(* IEC 61131-3 sources: s7-to-codesys/src/POUs/Lang/Converted/FB_BackwashGraph, 2 files *)

(* ---- FB_BackwashGraph.decl.st ---- *)
// Назначение: Промывка фильтра (GRAPH)
//             Промывка скорого фильтра (GRAPH S7-1500), шаги S1–S6. S1 Idle (начальный): N xReady.
//             T1 Start: xStart. S2 Drain: N xDrainValve, S xWashActive, событие S1 — iWashCount + 1;
//             контроль xValveFault держит шаг до квитирования ACK_EF (ERR_FLT = 1). После S2 альтернатива:
//             T2 LongWash (xLevelLow AND NOT xShortWash) — параллельно S3 Air (N xBlower, D xAirValve 2 с)
//             и S4 Rinse (NC xWashPump, блокировка xPumpOk), синхронизация T4 AirDone: Air.T >= 10 с;
//             T3 ShortWash (xLevelLow AND xShortWash) — S5 QuickRinse (N xWashPump), T5 QuickDone: xLevelHigh.
//             S6 Refill: N xInletValve, R xWashActive; T6 Full: xLevelHigh — прыжок к S1. Постоперация:
//             xValvesBusy := xDrainValve OR xInletValve. INIT_SQ — начальное состояние, OFF_SQ — шаги выключены.
// Автор:      WTP2 (исходный блок S7); перевод в ST — s7conv 0.1.0
// Версия:     0.1 (исходный блок S7)
// Документ:   docs/CONVERSION_REPORT.md, docs/MAPPING.md
// Источник:   samples/lang/FB_BackwashGraph.xml, GRAPH, SW.Blocks.FB "FB_BackwashGraph", пространство имён
//             Interface/v5, FAMILY Filters
// Сгенерировано s7conv: пометки MIGRATION-CHECK и MIGRATION-TODO требуют ручного разбора.
FUNCTION_BLOCK FB_BackwashGraph
VAR_INPUT
    OFF_SQ : BOOL;  // Выключить последовательность
    INIT_SQ : BOOL;  // Начальное состояние
    ACK_EF : BOOL;  // Квитирование ошибок контроля
    xStart : BOOL;  // Пуск промывки
    xLevelLow : BOOL;  // Уровень ниже сливного
    xLevelHigh : BOOL;  // Фильтр заполнен
    xShortWash : BOOL;  // Короткая промывка (без продувки)
    xPumpOk : BOOL := TRUE;  // Насос промывки исправен
    xValveFault : BOOL;  // Неисправность сливной задвижки
END_VAR
VAR_OUTPUT
    ERR_FLT : BOOL;  // Ошибка контроля (до квитирования)
    xReady : BOOL;  // Готов к промывке
    xDrainValve : BOOL;  // Сливная задвижка
    xBlower : BOOL;  // Воздуходувка
    xAirValve : BOOL;  // Задвижка воздуха
    xWashPump : BOOL;  // Насос промывки
    xInletValve : BOOL;  // Задвижка подачи
    xWashActive : BOOL;  // Промывка идёт
    xValvesBusy : BOOL;  // Задвижки в работе
    iWashCount : INT;  // Число промывок
END_VAR
VAR_TEMP
    tGraphNow : TIME;  // GRAPH: время вызова (F_S7Now)
    xIdle_Prev : BOOL;  // шаг S1: активен в прошлом вызове
    xIdle_S1 : BOOL;  // шаг S1: событие S1 (активирован)
    xIdle_S0 : BOOL;  // шаг S1: событие S0 (выключен)
    xDrain_Prev : BOOL;  // шаг S2: активен в прошлом вызове
    xDrain_S1 : BOOL;  // шаг S2: событие S1 (активирован)
    xDrain_S0 : BOOL;  // шаг S2: событие S0 (выключен)
    xAir_Prev : BOOL;  // шаг S3: активен в прошлом вызове
    xAir_S1 : BOOL;  // шаг S3: событие S1 (активирован)
    xAir_S0 : BOOL;  // шаг S3: событие S0 (выключен)
    xRinse_Prev : BOOL;  // шаг S4: активен в прошлом вызове
    xRinse_S1 : BOOL;  // шаг S4: событие S1 (активирован)
    xRinse_S0 : BOOL;  // шаг S4: событие S0 (выключен)
    xRinse_Il : BOOL;  // шаг S4: блокировка выполнена
    xQuickRinse_Prev : BOOL;  // шаг S5: активен в прошлом вызове
    xQuickRinse_S1 : BOOL;  // шаг S5: событие S1 (активирован)
    xQuickRinse_S0 : BOOL;  // шаг S5: событие S0 (выключен)
    xRefill_Prev : BOOL;  // шаг S6: активен в прошлом вызове
    xRefill_S1 : BOOL;  // шаг S6: событие S1 (активирован)
    xRefill_S0 : BOOL;  // шаг S6: событие S0 (выключен)
    xGraphHold : BOOL;  // GRAPH: INIT_SQ, OFF_SQ или первый вызов — переходы не срабатывают
    xT1_Cond : BOOL;  // переход T1 Start: условие
    xT1_Fire : BOOL;  // переход T1: срабатывает
    xT2_Cond : BOOL;  // переход T2 LongWash: условие
    xT2_Fire : BOOL;  // переход T2: срабатывает
    xT3_Cond : BOOL;  // переход T3 ShortWash: условие
    xT3_Fire : BOOL;  // переход T3: срабатывает
    xT4_Cond : BOOL;  // переход T4 AirDone: условие
    xT4_Fire : BOOL;  // переход T4: срабатывает
    xT5_Cond : BOOL;  // переход T5 QuickDone: условие
    xT5_Fire : BOOL;  // переход T5: срабатывает
    xT6_Cond : BOOL;  // переход T6 Full: условие
    xT6_Fire : BOOL;  // переход T6: срабатывает
    xDrain_Sv : BOOL;  // шаг S2: условие контроля
END_VAR
VAR
    GraphInitDone : BOOL;  // GRAPH: начальное состояние установлено
    Idle_X : BOOL;  // шаг S1 Idle активен
    Idle_T : TIME;  // шаг S1: время активности (последней)
    Idle_Start : TIME;  // шаг S1: момент активации
    Drain_X : BOOL;  // шаг S2 Drain активен
    Drain_T : TIME;  // шаг S2: время активности (последней)
    Drain_Start : TIME;  // шаг S2: момент активации
    Drain_SvErr : BOOL;  // шаг S2: ошибка контроля
    Air_X : BOOL;  // шаг S3 Air активен
    Air_T : TIME;  // шаг S3: время активности (последней)
    Air_Start : TIME;  // шаг S3: момент активации
    Rinse_X : BOOL;  // шаг S4 Rinse активен
    Rinse_T : TIME;  // шаг S4: время активности (последней)
    Rinse_Start : TIME;  // шаг S4: момент активации
    QuickRinse_X : BOOL;  // шаг S5 QuickRinse активен
    QuickRinse_T : TIME;  // шаг S5: время активности (последней)
    QuickRinse_Start : TIME;  // шаг S5: момент активации
    Refill_X : BOOL;  // шаг S6 Refill активен
    Refill_T : TIME;  // шаг S6: время активности (последней)
    Refill_Start : TIME;  // шаг S6: момент активации
END_VAR

(* ---- FB_BackwashGraph.impl.st ---- *)
// Сеть 1 (GRAPH): Промывка фильтра
tGraphNow := F_S7Now();
// Состояние шагов прошлого вызова: события S1/S0 — и от INIT_SQ, OFF_SQ
xIdle_Prev := Idle_X;
xDrain_Prev := Drain_X;
xAir_Prev := Air_X;
xRinse_Prev := Rinse_X;
xQuickRinse_Prev := QuickRinse_X;
xRefill_Prev := Refill_X;
xGraphHold := INIT_SQ OR NOT GraphInitDone OR OFF_SQ;
// Начальное состояние (INIT_SQ, первый вызов) и выключение (OFF_SQ)
IF INIT_SQ OR NOT GraphInitDone THEN
    GraphInitDone := TRUE;
    Idle_X := TRUE;
    Idle_Start := tGraphNow;
    Idle_T := T#0MS;
    Drain_X := FALSE;
    Air_X := FALSE;
    Rinse_X := FALSE;
    QuickRinse_X := FALSE;
    Refill_X := FALSE;
    Drain_SvErr := FALSE;
END_IF
IF OFF_SQ THEN
    Idle_X := FALSE;
    Drain_X := FALSE;
    Air_X := FALSE;
    Rinse_X := FALSE;
    QuickRinse_X := FALSE;
    Refill_X := FALSE;
END_IF
// Квитирование ошибок контроля (ACK_EF): в этом вызове переход возможен
IF ACK_EF THEN
    Drain_SvErr := FALSE;
END_IF
// Время активных шагов
IF Idle_X THEN
    Idle_T := F_S7TimeDiff(tGraphNow, Idle_Start);
END_IF
IF Drain_X THEN
    Drain_T := F_S7TimeDiff(tGraphNow, Drain_Start);
END_IF
IF Air_X THEN
    Air_T := F_S7TimeDiff(tGraphNow, Air_Start);
END_IF
IF Rinse_X THEN
    Rinse_T := F_S7TimeDiff(tGraphNow, Rinse_Start);
END_IF
IF QuickRinse_X THEN
    QuickRinse_T := F_S7TimeDiff(tGraphNow, QuickRinse_Start);
END_IF
IF Refill_X THEN
    Refill_T := F_S7TimeDiff(tGraphNow, Refill_Start);
END_IF
// Условия переходов (сети LAD/FBD)
// MIGRATION-CHECK: элемент «TrCoil»: имя и пины в SimaticML не подтверждены открытым экспортом
//                  (docs/MAPPING_LADFBD.md, уровень L) (FB_BackwashGraph.xml, сеть 1 (GRAPH), переход T1, UId 23)
xT1_Cond := xStart;
// MIGRATION-CHECK: элемент «TrCoil»: имя и пины в SimaticML не подтверждены открытым экспортом
//                  (docs/MAPPING_LADFBD.md, уровень L) (FB_BackwashGraph.xml, сеть 1 (GRAPH), переход T2, UId 25)
xT2_Cond := xLevelLow AND NOT xShortWash;
// MIGRATION-CHECK: элемент «TrCoil»: имя и пины в SimaticML не подтверждены открытым экспортом
//                  (docs/MAPPING_LADFBD.md, уровень L) (FB_BackwashGraph.xml, сеть 1 (GRAPH), переход T3, UId 25)
xT3_Cond := xLevelLow AND xShortWash;
// MIGRATION-CHECK: элемент «TrCoil»: имя и пины в SimaticML не подтверждены открытым экспортом
//                  (docs/MAPPING_LADFBD.md, уровень L) (FB_BackwashGraph.xml, сеть 1 (GRAPH), переход T4, UId 24)
xT4_Cond := Air_T >= T#10S;
// MIGRATION-CHECK: элемент «TrCoil»: имя и пины в SimaticML не подтверждены открытым экспортом
//                  (docs/MAPPING_LADFBD.md, уровень L) (FB_BackwashGraph.xml, сеть 1 (GRAPH), переход T5, UId 23)
xT5_Cond := xLevelHigh;
// MIGRATION-CHECK: элемент «TrCoil»: имя и пины в SimaticML не подтверждены открытым экспортом
//                  (docs/MAPPING_LADFBD.md, уровень L) (FB_BackwashGraph.xml, сеть 1 (GRAPH), переход T6, UId 23)
xT6_Cond := xLevelHigh;
// Срабатывание: предшественники активны, условие, нет ошибки контроля; альтернативы — слева направо
xT1_Fire := Idle_X AND xT1_Cond AND NOT xGraphHold;
xT2_Fire := Drain_X AND xT2_Cond AND NOT xGraphHold AND NOT Drain_SvErr;
// MIGRATION-CHECK: альтернативная ветвь: из одновременно истинных переходов срабатывает левый (первый); настройку
//                  блока S7-1500 сверить (FB_BackwashGraph.xml, сеть 1 (GRAPH), переход T3)
xT3_Fire := Drain_X AND xT3_Cond AND NOT xGraphHold AND NOT Drain_SvErr AND NOT xT2_Fire;
xT4_Fire := Air_X AND Rinse_X AND xT4_Cond AND NOT xGraphHold;
xT5_Fire := QuickRinse_X AND xT5_Cond AND NOT xGraphHold;
xT6_Fire := Refill_X AND xT6_Cond AND NOT xGraphHold;
// Переключение: сначала выключение предшественников, затем включение преемников
IF xT1_Fire THEN
    Idle_X := FALSE;
END_IF
IF xT2_Fire THEN
    Drain_X := FALSE;
END_IF
IF xT3_Fire THEN
    Drain_X := FALSE;
END_IF
IF xT4_Fire THEN
    Air_X := FALSE;
    Rinse_X := FALSE;
END_IF
IF xT5_Fire THEN
    QuickRinse_X := FALSE;
END_IF
IF xT6_Fire THEN
    Refill_X := FALSE;
END_IF
IF xT1_Fire THEN
    Drain_X := TRUE;
END_IF
IF xT2_Fire THEN
    Air_X := TRUE;
    Rinse_X := TRUE;
END_IF
IF xT3_Fire THEN
    QuickRinse_X := TRUE;
END_IF
IF xT4_Fire THEN
    Refill_X := TRUE;
END_IF
IF xT5_Fire THEN
    Refill_X := TRUE;
END_IF
IF xT6_Fire THEN
    Idle_X := TRUE;
END_IF
// События шагов S1/S0; активация — новый отсчёт времени
xIdle_S1 := Idle_X AND NOT xIdle_Prev;
xIdle_S0 := xIdle_Prev AND NOT Idle_X;
IF xIdle_S1 THEN
    Idle_Start := tGraphNow;
    Idle_T := T#0MS;
END_IF
xDrain_S1 := Drain_X AND NOT xDrain_Prev;
xDrain_S0 := xDrain_Prev AND NOT Drain_X;
IF xDrain_S1 THEN
    Drain_Start := tGraphNow;
    Drain_T := T#0MS;
END_IF
xAir_S1 := Air_X AND NOT xAir_Prev;
xAir_S0 := xAir_Prev AND NOT Air_X;
IF xAir_S1 THEN
    Air_Start := tGraphNow;
    Air_T := T#0MS;
END_IF
xRinse_S1 := Rinse_X AND NOT xRinse_Prev;
xRinse_S0 := xRinse_Prev AND NOT Rinse_X;
IF xRinse_S1 THEN
    Rinse_Start := tGraphNow;
    Rinse_T := T#0MS;
END_IF
xQuickRinse_S1 := QuickRinse_X AND NOT xQuickRinse_Prev;
xQuickRinse_S0 := xQuickRinse_Prev AND NOT QuickRinse_X;
IF xQuickRinse_S1 THEN
    QuickRinse_Start := tGraphNow;
    QuickRinse_T := T#0MS;
END_IF
xRefill_S1 := Refill_X AND NOT xRefill_Prev;
xRefill_S0 := xRefill_Prev AND NOT Refill_X;
IF xRefill_S1 THEN
    Refill_Start := tGraphNow;
    Refill_T := T#0MS;
END_IF
// Контроль шага S2 Drain
// MIGRATION-CHECK: элемент «SvCoil»: имя и пины в SimaticML не подтверждены открытым экспортом
//                  (docs/MAPPING_LADFBD.md, уровень L) (FB_BackwashGraph.xml, сеть 1 (GRAPH), шаг S2, контроль, UId
//                  23)
xDrain_Sv := xValveFault;
// MIGRATION-CHECK: контроль S2: ошибка защёлкивается и держит шаг до ACK_EF; Si.U и сообщения ProDiag не
//                  переносятся (FB_BackwashGraph.xml, сеть 1 (GRAPH), шаг S2, контроль)
IF Drain_X AND xDrain_Sv THEN
    Drain_SvErr := TRUE;
END_IF
// Блокировка шага S4 Rinse
// MIGRATION-CHECK: элемент «IlCoil»: имя и пины в SimaticML не подтверждены открытым экспортом
//                  (docs/MAPPING_LADFBD.md, уровень L) (FB_BackwashGraph.xml, сеть 1 (GRAPH), шаг S4, блокировка,
//                  UId 23)
xRinse_Il := xPumpOk;
// Действия шага S1 Idle
IF Idle_X OR xIdle_S0 THEN
    xReady := Idle_X;
END_IF
// Действия шага S2 Drain
IF Drain_X OR xDrain_S0 THEN
    xDrainValve := Drain_X;
END_IF
IF Drain_X THEN
    xWashActive := TRUE;
END_IF
IF xDrain_S1 THEN
    iWashCount := iWashCount + 1;
END_IF
// Действия шага S3 Air
IF Air_X OR xAir_S0 THEN
    xBlower := Air_X;
END_IF
// MIGRATION-CHECK: S3: D #xAirValve, T#2S — по времени шага #Air_T (F_S7Now); в SFC — IEC D по своему таймеру
//                  (FB_BackwashGraph.xml, сеть 1 (GRAPH), шаг S3, действие 2)
IF Air_X OR xAir_S0 THEN
    xAirValve := Air_X AND Air_T >= T#2S;
END_IF
// Действия шага S4 Rinse
IF Rinse_X OR xRinse_S0 THEN
    xWashPump := Rinse_X AND xRinse_Il;
END_IF
// Действия шага S5 QuickRinse
IF QuickRinse_X OR xQuickRinse_S0 THEN
    xWashPump := QuickRinse_X;
END_IF
// Действия шага S6 Refill
IF Refill_X OR xRefill_S0 THEN
    xInletValve := Refill_X;
END_IF
IF Refill_X THEN
    xWashActive := FALSE;
END_IF
ERR_FLT := Drain_SvErr;
// Постоперация 1
xValvesBusy := xDrainValve OR xInletValve;
